{region 'Documentation'}
(*!
<summary>Checks inequality with the forbidden LWORD value.</summary>
*)
{endregion}
FUNCTION_BLOCK AssertNotEqual_LWord EXTENDS AssertionBase
VAR_INPUT
    IN : LWORD; //! Actual value checked or observed by this Assertion.
    Expected : LWORD; //! Value that must differ from IN under this Assertion's comparison rules.
END_VAR

SUPER^();

{region 'Documentation'}
(*!
<summary>Check inequality with the forbidden LWORD value.</summary>
*)
{endregion}
METHOD PROTECTED Assert
VAR
    Message : STRING(GVL_Constants.MessageLength);
    ExpectedText : STRING(GVL_Constants.AssertionValueLength);
    ActualText : STRING(GVL_Constants.AssertionValueLength);
END_VAR
VAR CONSTANT
    HexDigitCount : USINT := 16;
END_VAR
IF NOT EvaluationActive THEN
    RETURN;
END_IF;

IF Result = E_Result.Error THEN
    RETURN;
END_IF;

IF Result = E_Result.Failed THEN
    RETURN;
END_IF;

IF IN = Expected THEN
    ExpectedText := CreateAssertionTextValue_Hex(Value := Expected,
        DigitCount := HexDigitCount);
    ActualText := CreateAssertionTextValue_Hex(Value := IN,
        DigitCount := HexDigitCount);
    Message := CONCAT('Assertion failed: values are equal but should differ. NotExpected = ',
        ExpectedText);
    Message := CONCAT(Message, ', Actual = ');
    Message := CONCAT(Message, ActualText);
    Message := CONCAT(Message, '.');
    Fail(Message := Message);
    RETURN;
END_IF;

Pass();
END_METHOD

END_FUNCTION_BLOCK

(* stored: Version 1.1.0.1
   POU AssertNotEqual_LWord: Id {a5feabd9-a50f-42d9-9657-bd9558f43faa}, SpecialFunc None
   Folder Internal: Id {bd686b57-a176-4125-9841-0999d41ec78f}
   Method Assert: Id {83c2a303-0e45-4524-926d-a5073f7e4963} *)
